// TIA Portal V21 program export: 0 tag tables, 0 data types, 0 data blocks, 2 code blocks (in call order from the OBs), 0 instance data blocks

ORGANIZATION_BLOCK "LongNames"   // OB1, LAD
BEGIN

REGION Network 1: Long tag names
   // A comment that runs on.
   // And a second line.
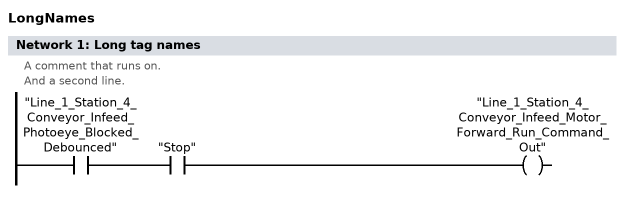
   RUNG wire#powerrail
      Contact( "Line_1_Station_4_Conveyor_Infeed_Photoeye_Blocked_Debounced" )
      Contact( "Stop" )
      Coil( "Line_1_Station_4_Conveyor_Infeed_Motor_Forward_Run_Command_Out" )
   END_RUNG
   // the same network as SCL:
   "Line_1_Station_4_Conveyor_Infeed_Motor_Forward_Run_Command_Out" := "Line_1_Station_4_Conveyor_Infeed_Photoeye_Blocked_Debounced" AND "Stop";
END_REGION
END_ORGANIZATION_BLOCK

FUNCTION_BLOCK "Mixed"   // FB1, LAD
BEGIN

REGION Network 1: Unknown part
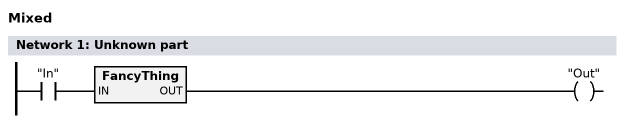
   // no SCL statement known for FancyThing: written as a call
   "Out" := FancyThing("In");
END_REGION

REGION Network 2 (SCL): SCL inside
END_REGION

REGION Network 3: Empty
END_REGION
END_FUNCTION_BLOCK
